Fanuc KAREL source: kt00134.KL

-- PROVISIONAL review KL for V1013-1; original PC SHA256 e7f9434cd711eb99100168121dec9bbb380e72e088285b8ad1c215996fd69cc3
-- Incomplete behavior may be omitted. Consult companion uncertainty JSON. Do not deploy.
PROGRAM KT00134
%NOLOCKGROUP
VAR
  I1 : INTEGER
  OUT : REAL
-- UNRESOLVED_DECL Y2 type=002018
BEGIN
  -- UNRESOLVED_PC offsets 5-16; opcodes 2E,23
  -- UNRESOLVED_PC offsets 21-35; opcodes 2E,22,9D,33,B2
  -- UNRESOLVED_PC offsets 40-63; opcodes 21,22,9D,33,B1,55,64,23
  -- UNRESOLVED_PC offsets 68-72; opcodes 7F
END KT00134
